# EPICS substitutions: db/Festo/ecmcFesto-CMMT-ST.substitutions
file "ecmcFesto-CMMT-ST.template" { pattern
  { CH_ID }
  { 01    }
}

file "ecmcFesto-CMMT-ST_Enc-chX.template" { pattern
  { CH_ID }
  { 01    }
  { 02    }
}

file "ecmcFesto-CMMT-ST_Enc.template" { pattern
  { CH_ID }
  { X     }
}

# ecmcDS402Enable
file "ecmcDS402Enable-chX.template"
{
  pattern {CH_ID}
          {01   }
}
